FUNCTION_BLOCK FB_Valve
var_input
R:bool;
nSpeed:int; // speed
end_var
VAR
sTimer:TON;
sbDone : BOOL;
END_VAR

if R then
sTimer(IN:=TRUE,PT:=T#5S,Q=>sbDone);
end_if

METHOD M_Reset : BOOL
VAR_INPUT
bForce:BOOL;
END_VAR
VAR
x : INT;
END_VAR
x:=0;
M_Reset:=TRUE;
END_METHOD

END_FUNCTION_BLOCK

(* stored: Version 1.1.0.1, ProductVersion 3.1.4024.12
   POU FB_Valve: Id {11111111-2222-3333-4444-555555555555}, SpecialFunc None
   Method M_Reset: Id {aaaaaaaa-2222-3333-4444-555555555555} *)
